Fanuc KAREL source: kd00053.KL

-- PROVISIONAL review KL for V770-1; original PC SHA256 6663f1f33fc36c0b7cd47bc32af10c3a004f0117a154e5a205052fcff9fa217b
-- Incomplete behavior may be omitted. Consult companion uncertainty JSON. Do not deploy.
PROGRAM KD00053
%NOLOCKGROUP
VAR
  I : INTEGER
  J : INTEGER
  B : BOOLEAN
  R : REAL
  S : STRING[80]
BEGIN
  -- UNRESOLVED_PC offsets 5-19; opcodes 21,9D,52,23
  -- UNRESOLVED_PC offsets 24-28; opcodes 7F
END KD00053
